(* IEC 61131-3 sources: model-first-plc-agent-ai/results/T3-W-20, 2 files *)

(* ---- a1_code.st ---- *)
FUNCTION_BLOCK FillingRuntime
VAR_INPUT
    start : BOOL;
    stop : BOOL;
    LSH : BOOL;
    LSHH : BOOL;
    TON_Duration : TIME;
    TOF_Duration : TIME;
END_VAR
VAR_OUTPUT
    fill_valve : BOOL;
    discharge_valve : BOOL;
END_VAR
VAR
    x0 : BOOL := TRUE;
    x1 : BOOL := FALSE;
    x2 : BOOL := FALSE;
    t1 : BOOL;
    t2 : BOOL;
    t3 : BOOL;
    t4 : BOOL;
    t5 : BOOL;
    ton_q : BOOL;
    tof_q : BOOL;
    FillingTimer : TON;
    PauseTimer : TOF;
END_VAR

(* Both timers are evaluated every scan using filling-step activity. *)
FillingTimer(IN := x1, PT := TON_Duration);
PauseTimer(IN := x1, PT := TOF_Duration);

ton_q := FillingTimer.Q;
tof_q := PauseTimer.Q;

(* Evaluate all transitions against the same current situation. *)
t1 := x0 AND start AND NOT stop AND NOT LSH AND NOT LSHH;
t2 := x1 AND ton_q AND NOT stop AND NOT LSH AND NOT LSHH;
t3 := x2 AND NOT tof_q AND NOT stop AND NOT LSH AND NOT LSHH;
t4 := x1 AND (stop OR LSH OR LSHH);
t5 := x2 AND (stop OR LSH OR LSHH);

(* Apply the simultaneous situation update. *)
x0 := (x0 AND NOT t1) OR t4 OR t5;
x1 := (x1 AND NOT (t2 OR t4)) OR t1 OR t3;
x2 := (x2 AND NOT (t3 OR t5)) OR t2;

(* Continuous, non-stored actions. *)
fill_valve := x1;
discharge_valve := FALSE;

END_FUNCTION_BLOCK

PROGRAM Main
VAR
    StartCommand AT %IX100.0 : BOOL;
    StopCommand AT %IX100.1 : BOOL;
    LSH AT %IX100.2 : BOOL;
    LSHH AT %IX100.3 : BOOL;
    FillValve AT %QX100.0 : BOOL;
    DischargeValve AT %QX100.1 : BOOL;
END_VAR
VAR
    (* Configurable example presets; set to the required process values. *)
    TON_Duration : TIME := T#5s;
    TOF_Duration : TIME := T#5s;
    StartEdge : R_TRIG;
    Controller : FillingRuntime;
END_VAR

StartEdge(CLK := StartCommand);

Controller(
    start := StartEdge.Q,
    stop := StopCommand,
    LSH := LSH,
    LSHH := LSHH,
    TON_Duration := TON_Duration,
    TOF_Duration := TOF_Duration
);

FillValve := Controller.fill_valve;
DischargeValve := Controller.discharge_valve;

END_PROGRAM

(* ---- a2_code.st ---- *)
FUNCTION_BLOCK FB_TankFilling
VAR_INPUT
    StartCommand : BOOL;
    StopCommand : BOOL;
    LSH : BOOL;
    LSHH : BOOL;
    TON_Duration : TIME;
    TOF_Duration : TIME;
END_VAR
VAR_OUTPUT
    fill_valve : BOOL;
    discharge_valve : BOOL;
END_VAR
VAR
    cycle_state : INT := 0;
    start_edge : R_TRIG;
    filling_timer : TON;
    pause_timer : TOF;
    start : BOOL;
    stop : BOOL;
    ton_q : BOOL;
    tof_q : BOOL;
    filling_active : BOOL;
END_VAR

start_edge(CLK := StartCommand);
start := start_edge.Q;
stop := StopCommand;

(* Both timers measure the activity of the filling step. *)
filling_active := (cycle_state = 1);
filling_timer(IN := filling_active, PT := TON_Duration);
pause_timer(IN := filling_active, PT := TOF_Duration);

ton_q := filling_timer.Q;
tof_q := pause_timer.Q;

(* Stop has priority over all normal transitions. *)
IF stop THEN
    cycle_state := 0;
ELSE
    CASE cycle_state OF
        0:
            IF start AND NOT LSH THEN
                cycle_state := 1;
            END_IF;

        1:
            IF LSH THEN
                cycle_state := 0;
            ELSIF ton_q THEN
                cycle_state := 2;
            END_IF;

        2:
            IF LSH THEN
                cycle_state := 0;
            ELSIF NOT tof_q THEN
                cycle_state := 1;
            END_IF;

        ELSE
            cycle_state := 0;
    END_CASE;
END_IF;

(* LSHH is monitored by the plant; no additional transition is specified. *)
fill_valve := (cycle_state = 1) AND NOT stop;
discharge_valve := FALSE;

END_FUNCTION_BLOCK

PROGRAM Main
VAR
    StartCommand AT %IX100.0 : BOOL;
    StopCommand AT %IX100.1 : BOOL;
    LSH AT %IX100.2 : BOOL;
    LSHH AT %IX100.3 : BOOL;
    FillValve AT %QX100.0 : BOOL;
    DischargeValve AT %QX100.1 : BOOL;
END_VAR
VAR
    tank_controller : FB_TankFilling;
    (* Example presets; configure these for the required cycle timing. *)
    TON_Duration : TIME := T#5s;
    TOF_Duration : TIME := T#3s;
END_VAR

tank_controller(
    StartCommand := StartCommand,
    StopCommand := StopCommand,
    LSH := LSH,
    LSHH := LSHH,
    TON_Duration := TON_Duration,
    TOF_Duration := TOF_Duration
);

FillValve := tank_controller.fill_valve;
DischargeValve := tank_controller.discharge_valve;

END_PROGRAM
